(* IEC 61131-3 sources: trust-platform/examples/OSCAT/pasteurizer_quality_chain/oop/src, 3 files *)

(* ---- Main.st ---- *)
(* Record role: PasteurizerResult is a deterministic PLC-side record for tests and runtime readers. *)
TYPE PasteurizerResult :
STRUCT
    ForwardDivert : BOOL;
    DivertToRecirc : BOOL;
    RequiredTemperature : REAL;
    RequiredHoldSeconds : INT;
    SequenceStep : INT;
END_STRUCT
END_TYPE

(* Record role: QualityAlarmEvent is a deterministic PLC-side record for tests and runtime readers. *)
TYPE QualityAlarmEvent :
STRUCT
    TemperatureC : REAL;
    FlowRateLpm : REAL;
    RequiredTemperatureC : REAL;
    OperatorAck : BOOL;
    SupervisorOnline : BOOL;
END_STRUCT
END_TYPE

(* Pattern role: IQualityAlarmHandler is the contract boundary for the Chain of Responsibility and Template Method example. *)
INTERFACE IQualityAlarmHandler
    METHOD SetNext
    VAR_INPUT
        NextHandler : IQualityAlarmHandler;
    END_VAR
    END_METHOD

    METHOD Handle : BOOL
    VAR_INPUT
        Event : QualityAlarmEvent;
    END_VAR
    END_METHOD

    PROPERTY HandlerId : INT
    GET
    END_GET
    END_PROPERTY
END_INTERFACE

(* Composition role: BasePasteurizerTemplate owns the collaborating objects used by this Chain of Responsibility and Template Method example. *)
FUNCTION_BLOCK BasePasteurizerTemplate
VAR
    TempFilter : Pt2Filter;
    DivertCounter : DwordCounter;
    LastResult : PasteurizerResult;
END_VAR

METHOD PUBLIC Initialize
TempFilter.Initialize();
TempFilter.Configure(TimeConstant := T#1s, Damping := REAL#1.0, Gain := REAL#1.0);
DivertCounter.Initialize();
DivertCounter.Configure(StepSize := DWORD#1, MaxValue := DWORD#16#FFFFFFFF);
END_METHOD

METHOD PUBLIC RequiredTemperature : REAL
RequiredTemperature := REAL#72.0;
END_METHOD

METHOD PUBLIC RequiredHoldSeconds : INT
RequiredHoldSeconds := INT#15;
END_METHOD

METHOD PUBLIC Preheat : BOOL
VAR_INPUT
    ProductPresent : BOOL;
END_VAR
Preheat := ProductPresent;
END_METHOD

METHOD PUBLIC Heat : BOOL
VAR_INPUT
    ProductTemp : REAL;
END_VAR
Heat := ProductTemp >= RequiredTemperature();
END_METHOD

METHOD PUBLIC Hold : BOOL
VAR_INPUT
    HoldSeconds : INT;
END_VAR
Hold := HoldSeconds >= RequiredHoldSeconds();
END_METHOD

METHOD PUBLIC Chill : BOOL
VAR_INPUT
    FlowRate : REAL;
END_VAR
Chill := FlowRate >= REAL#100.0;
END_METHOD

METHOD PUBLIC RouteProduct : BOOL
VAR_INPUT
    HeatOk : BOOL;
    HoldOk : BOOL;
    ChillOk : BOOL;
END_VAR
RouteProduct := HeatOk AND HoldOk AND ChillOk;
END_METHOD

METHOD PUBLIC RunTemplate : PasteurizerResult
VAR_INPUT
    ProductPresent : BOOL;
    ProductTemp : REAL;
    FlowRate : REAL;
    HoldSeconds : INT;
END_VAR
VAR
    HeatOk : BOOL;
    HoldOk : BOOL;
    ChillOk : BOOL;
END_VAR
LastResult.RequiredTemperature := RequiredTemperature();
LastResult.RequiredHoldSeconds := RequiredHoldSeconds();
(* SequenceStep legend: 10=preheat wait, 20=heat, 40=recirculate/divert, 50=forward product. *)
IF NOT Preheat(ProductPresent := ProductPresent) THEN
    LastResult.SequenceStep := INT#10;
    LastResult.ForwardDivert := FALSE;
ELSIF NOT Heat(ProductTemp := ProductTemp) THEN
    LastResult.SequenceStep := INT#20;
    LastResult.ForwardDivert := FALSE;
ELSE
    HeatOk := TRUE;
    HoldOk := Hold(HoldSeconds := HoldSeconds);
    ChillOk := Chill(FlowRate := FlowRate);
    LastResult.ForwardDivert := RouteProduct(HeatOk := HeatOk, HoldOk := HoldOk, ChillOk := ChillOk);
    IF LastResult.ForwardDivert THEN
        LastResult.SequenceStep := INT#50;
    ELSE
        LastResult.SequenceStep := INT#40;
    END_IF;
END_IF;
LastResult.DivertToRecirc := NOT LastResult.ForwardDivert;
(* DwordCounter wraps COUNT_DR (edge-triggered: UP AND NOT LastUp).
   Drop the UP edge first so consecutive divert batches each generate
   a fresh rising edge and actually increment. *)
DivertCounter.Update(Up := FALSE, Down := FALSE);
IF LastResult.DivertToRecirc THEN
    DivertCounter.Update(Up := TRUE, Down := FALSE);
END_IF;
RunTemplate := LastResult;
END_METHOD
END_FUNCTION_BLOCK

(* Pattern role: MilkPasteurizer customizes inherited behavior in the Chain of Responsibility and Template Method example. *)
FUNCTION_BLOCK MilkPasteurizer EXTENDS BasePasteurizerTemplate
METHOD PUBLIC RequiredTemperature : REAL
RequiredTemperature := REAL#72.0;
END_METHOD

METHOD PUBLIC RequiredHoldSeconds : INT
RequiredHoldSeconds := INT#15;
END_METHOD
END_FUNCTION_BLOCK

(* Pattern role: CreamPasteurizer customizes inherited behavior in the Chain of Responsibility and Template Method example. *)
FUNCTION_BLOCK CreamPasteurizer EXTENDS BasePasteurizerTemplate
METHOD PUBLIC RequiredTemperature : REAL
RequiredTemperature := REAL#75.0;
END_METHOD

METHOD PUBLIC RequiredHoldSeconds : INT
RequiredHoldSeconds := INT#20;
END_METHOD
END_FUNCTION_BLOCK

(* Pattern role: LocalRecoveryHandler is a concrete implementation in the Chain of Responsibility and Template Method example. *)
FUNCTION_BLOCK LocalRecoveryHandler IMPLEMENTS IQualityAlarmHandler
VAR
    Next : IQualityAlarmHandler;
    HandlerIdValue : INT := INT#1;
    RecoveredValue : BOOL;
END_VAR

METHOD PUBLIC SetNext
VAR_INPUT
    NextHandler : IQualityAlarmHandler;
END_VAR
Next := NextHandler;
END_METHOD

METHOD PUBLIC Handle : BOOL
VAR_INPUT
    Event : QualityAlarmEvent;
END_VAR
(* Reset on entry so the flag reflects only the current event. *)
RecoveredValue := FALSE;
IF (Event.TemperatureC >= (Event.RequiredTemperatureC - REAL#1.0)) AND (Event.FlowRateLpm >= REAL#100.0) THEN
    RecoveredValue := TRUE;
    Handle := TRUE;
ELSE
    Handle := Next.Handle(Event := Event);
END_IF;
END_METHOD

METHOD PUBLIC ResetFlag
RecoveredValue := FALSE;
END_METHOD

PUBLIC PROPERTY HandlerId : INT
GET
    HandlerId := HandlerIdValue;
END_GET
END_PROPERTY

PUBLIC PROPERTY Recovered : BOOL
GET
    Recovered := RecoveredValue;
END_GET
END_PROPERTY
END_FUNCTION_BLOCK

(* Pattern role: OperatorAcknowledgeHandler is a concrete implementation in the Chain of Responsibility and Template Method example. *)
FUNCTION_BLOCK OperatorAcknowledgeHandler IMPLEMENTS IQualityAlarmHandler
VAR
    Next : IQualityAlarmHandler;
    HandlerIdValue : INT := INT#2;
    AcknowledgedValue : BOOL;
END_VAR

METHOD PUBLIC SetNext
VAR_INPUT
    NextHandler : IQualityAlarmHandler;
END_VAR
Next := NextHandler;
END_METHOD

METHOD PUBLIC Handle : BOOL
VAR_INPUT
    Event : QualityAlarmEvent;
END_VAR
(* Reset on entry so the flag reflects only the current event. *)
AcknowledgedValue := FALSE;
IF Event.OperatorAck THEN
    AcknowledgedValue := TRUE;
    Handle := TRUE;
ELSE
    Handle := Next.Handle(Event := Event);
END_IF;
END_METHOD

METHOD PUBLIC ResetFlag
AcknowledgedValue := FALSE;
END_METHOD

PUBLIC PROPERTY HandlerId : INT
GET
    HandlerId := HandlerIdValue;
END_GET
END_PROPERTY

PUBLIC PROPERTY Acknowledged : BOOL
GET
    Acknowledged := AcknowledgedValue;
END_GET
END_PROPERTY
END_FUNCTION_BLOCK

(* Pattern role: SupervisorEscalateHandler is a concrete implementation in the Chain of Responsibility and Template Method example. *)
FUNCTION_BLOCK SupervisorEscalateHandler IMPLEMENTS IQualityAlarmHandler
VAR
    Next : IQualityAlarmHandler;
    HandlerIdValue : INT := INT#3;
    EscalatedValue : BOOL;
END_VAR

METHOD PUBLIC SetNext
VAR_INPUT
    NextHandler : IQualityAlarmHandler;
END_VAR
Next := NextHandler;
END_METHOD

METHOD PUBLIC Handle : BOOL
VAR_INPUT
    Event : QualityAlarmEvent;
END_VAR
(* Reset on entry so the flag reflects only the current event. *)
EscalatedValue := FALSE;
IF Event.SupervisorOnline THEN
    EscalatedValue := TRUE;
    Handle := TRUE;
ELSE
    Handle := Next.Handle(Event := Event);
END_IF;
END_METHOD

METHOD PUBLIC ResetFlag
EscalatedValue := FALSE;
END_METHOD

PUBLIC PROPERTY HandlerId : INT
GET
    HandlerId := HandlerIdValue;
END_GET
END_PROPERTY

PUBLIC PROPERTY Escalated : BOOL
GET
    Escalated := EscalatedValue;
END_GET
END_PROPERTY
END_FUNCTION_BLOCK

(* Pattern role: BatchAbortHandler is a concrete implementation in the Chain of Responsibility and Template Method example. *)
FUNCTION_BLOCK BatchAbortHandler IMPLEMENTS IQualityAlarmHandler
VAR
    HandlerIdValue : INT := INT#4;
    AbortedValue : BOOL;
END_VAR

METHOD PUBLIC SetNext
VAR_INPUT
    NextHandler : IQualityAlarmHandler;
END_VAR
END_METHOD

METHOD PUBLIC Handle : BOOL
VAR_INPUT
    Event : QualityAlarmEvent;
END_VAR
(* Last handler in chain: always handles. Flag is set fresh each call. *)
AbortedValue := TRUE;
Handle := TRUE;
END_METHOD

METHOD PUBLIC ResetFlag
AbortedValue := FALSE;
END_METHOD

PUBLIC PROPERTY HandlerId : INT
GET
    HandlerId := HandlerIdValue;
END_GET
END_PROPERTY

PUBLIC PROPERTY Aborted : BOOL
GET
    Aborted := AbortedValue;
END_GET
END_PROPERTY
END_FUNCTION_BLOCK

(* Composition role: PasteurizerController owns the collaborating objects used by this Chain of Responsibility and Template Method example. *)
FUNCTION_BLOCK PasteurizerController
VAR
    Milk : MilkPasteurizer;
    Cream : CreamPasteurizer;
    Local : LocalRecoveryHandler;
    Operator : OperatorAcknowledgeHandler;
    Supervisor : SupervisorEscalateHandler;
    Abort : BatchAbortHandler;
    AlarmChain : IQualityAlarmHandler;
    LastResultValue : PasteurizerResult;
    LastHandlerIdValue : INT;
END_VAR

METHOD PUBLIC Initialize
Milk.Initialize();
Cream.Initialize();
Local.SetNext(NextHandler := Operator);
Operator.SetNext(NextHandler := Supervisor);
Supervisor.SetNext(NextHandler := Abort);
AlarmChain := Local;
END_METHOD

METHOD PUBLIC Update : PasteurizerResult
VAR_INPUT
    RecipeId : INT;
    ProductTemp : REAL;
    FlowRate : REAL;
    HoldSeconds : INT;
    OperatorAck : BOOL;
    SupervisorOnline : BOOL;
END_VAR
VAR
    Event : QualityAlarmEvent;
END_VAR
(* Clear cross-batch sticky state so LastHandlerId reflects only the current batch. *)
LastHandlerIdValue := INT#0;
Local.ResetFlag();
Operator.ResetFlag();
Supervisor.ResetFlag();
Abort.ResetFlag();
IF RecipeId = INT#2 THEN
    LastResultValue := Cream.RunTemplate(ProductPresent := TRUE, ProductTemp := ProductTemp, FlowRate := FlowRate, HoldSeconds := HoldSeconds);
ELSE
    LastResultValue := Milk.RunTemplate(ProductPresent := TRUE, ProductTemp := ProductTemp, FlowRate := FlowRate, HoldSeconds := HoldSeconds);
END_IF;

IF LastResultValue.DivertToRecirc THEN
    Event.TemperatureC := ProductTemp;
    Event.FlowRateLpm := FlowRate;
    Event.RequiredTemperatureC := LastResultValue.RequiredTemperature;
    Event.OperatorAck := OperatorAck;
    Event.SupervisorOnline := SupervisorOnline;
    AlarmChain.Handle(Event := Event);
    IF Abort.Aborted THEN
        LastHandlerIdValue := Abort.HandlerId;
    ELSIF Supervisor.Escalated THEN
        LastHandlerIdValue := Supervisor.HandlerId;
    ELSIF Operator.Acknowledged THEN
        LastHandlerIdValue := Operator.HandlerId;
    ELSIF Local.Recovered THEN
        LastHandlerIdValue := Local.HandlerId;
    END_IF;
END_IF;
Update := LastResultValue;
END_METHOD

PUBLIC PROPERTY ForwardDivert : BOOL
GET
    ForwardDivert := LastResultValue.ForwardDivert;
END_GET
END_PROPERTY

PUBLIC PROPERTY BatchAborted : BOOL
GET
    BatchAborted := Abort.Aborted;
END_GET
END_PROPERTY

PUBLIC PROPERTY LastHandlerId : INT
GET
    LastHandlerId := LastHandlerIdValue;
END_GET
END_PROPERTY

PUBLIC PROPERTY RequiredTemperature : REAL
GET
    RequiredTemperature := LastResultValue.RequiredTemperature;
END_GET
END_PROPERTY
END_FUNCTION_BLOCK

(* Scan role: Main wires the example objects and exposes the PLC call path under test. *)
PROGRAM Main
VAR
    Pasteurizer : PasteurizerController;
    RecipeId : INT;
    ProductTempRaw : INT;
    FlowRateRaw : INT;
    OperatorAck : BOOL;
    SupervisorOnline : BOOL;
    Result : PasteurizerResult;
    ForwardValveOut : BOOL;
    DivertValveOut : BOOL;
    AlarmOut : BOOL;
END_VAR

Pasteurizer.Initialize();
Result := Pasteurizer.Update(RecipeId := RecipeId, ProductTemp := INT_TO_REAL(ProductTempRaw), FlowRate := INT_TO_REAL(FlowRateRaw), HoldSeconds := INT#15, OperatorAck := OperatorAck, SupervisorOnline := SupervisorOnline);
ForwardValveOut := Result.ForwardDivert;
DivertValveOut := Result.DivertToRecirc;
AlarmOut := Result.DivertToRecirc;
END_PROGRAM

(* ---- Configuration.st ---- *)
CONFIGURATION PasteurizerQualityChainOopConfiguration
RESOURCE Cpu0 ON PLC
    TASK MainTask (INTERVAL := T#100ms, PRIORITY := 1);
    PROGRAM Pasteurizer WITH MainTask : Main;
END_RESOURCE
VAR_CONFIG
    Pasteurizer.RecipeId AT %IW0 : INT;
    Pasteurizer.ProductTempRaw AT %IW2 : INT;
    Pasteurizer.FlowRateRaw AT %IW4 : INT;
    Pasteurizer.OperatorAck AT %IX0.0 : BOOL;
    Pasteurizer.SupervisorOnline AT %IX0.1 : BOOL;
    Pasteurizer.ForwardValveOut AT %QX0.0 : BOOL;
    Pasteurizer.DivertValveOut AT %QX0.1 : BOOL;
    Pasteurizer.AlarmOut AT %QX0.2 : BOOL;
END_VAR
END_CONFIGURATION

(* ---- Tests.st ---- *)
TEST_PROGRAM PasteurizerTemplateUsesRecipeHooks
VAR
    Milk : MilkPasteurizer;
    Cream : CreamPasteurizer;
    MilkResult : PasteurizerResult;
    CreamResult : PasteurizerResult;
END_VAR

Milk.Initialize();
Cream.Initialize();
MilkResult := Milk.RunTemplate(ProductPresent := TRUE, ProductTemp := REAL#73.0, FlowRate := REAL#120.0, HoldSeconds := INT#15);
CreamResult := Cream.RunTemplate(ProductPresent := TRUE, ProductTemp := REAL#73.0, FlowRate := REAL#120.0, HoldSeconds := INT#15);
ASSERT_TRUE(IN := MilkResult.ForwardDivert);
ASSERT_FALSE(IN := CreamResult.ForwardDivert);
ASSERT_NEAR(EXPECTED := REAL#75.0, ACTUAL := CreamResult.RequiredTemperature, DELTA := REAL#0.001);
ASSERT_EQUAL(EXPECTED := INT#20, ACTUAL := CreamResult.RequiredHoldSeconds);
END_TEST_PROGRAM

TEST_PROGRAM QualityAlarmChainEscalatesToAbortWhenUnhandled
VAR
    Controller : PasteurizerController;
    Result : PasteurizerResult;
END_VAR

Controller.Initialize();
Result := Controller.Update(RecipeId := INT#1, ProductTemp := REAL#68.0, FlowRate := REAL#90.0, HoldSeconds := INT#5, OperatorAck := FALSE, SupervisorOnline := FALSE);
ASSERT_FALSE(IN := Result.ForwardDivert);
ASSERT_TRUE(IN := Controller.BatchAborted);
ASSERT_EQUAL(EXPECTED := INT#4, ACTUAL := Controller.LastHandlerId);
END_TEST_PROGRAM

TEST_PROGRAM QualityAlarmChainStopsAtOperatorAcknowledge
VAR
    Controller : PasteurizerController;
    Result : PasteurizerResult;
END_VAR

Controller.Initialize();
Result := Controller.Update(RecipeId := INT#1, ProductTemp := REAL#68.0, FlowRate := REAL#90.0, HoldSeconds := INT#5, OperatorAck := TRUE, SupervisorOnline := FALSE);
ASSERT_FALSE(IN := Result.ForwardDivert);
ASSERT_FALSE(IN := Controller.BatchAborted);
ASSERT_EQUAL(EXPECTED := INT#2, ACTUAL := Controller.LastHandlerId);
END_TEST_PROGRAM

(* Multi-batch chain regression: drives several different batches
   through one Controller. Catches the same bug class as
   tunnel_washer_chain — handler flags or LastHandlerId leaking
   between events because handlers don't reset their per-call state. *)
TEST_PROGRAM PasteurizerChainHandlesMultipleBatchesIndependently
VAR
    Controller : PasteurizerController;
    Result : PasteurizerResult;
END_VAR

Controller.Initialize();

(* Batch 1: bad temp + supervisor online -> escalates to supervisor (3) *)
Result := Controller.Update(RecipeId := INT#1, ProductTemp := REAL#68.0, FlowRate := REAL#90.0, HoldSeconds := INT#5, OperatorAck := FALSE, SupervisorOnline := TRUE);
ASSERT_EQUAL(EXPECTED := INT#3, ACTUAL := Controller.LastHandlerId);

(* Batch 2: same bad temp but operator now acks -> stops at handler 2.
   LastHandlerId must reflect the new outcome, not the previous (3). *)
Result := Controller.Update(RecipeId := INT#1, ProductTemp := REAL#68.0, FlowRate := REAL#90.0, HoldSeconds := INT#5, OperatorAck := TRUE, SupervisorOnline := FALSE);
ASSERT_EQUAL(EXPECTED := INT#2, ACTUAL := Controller.LastHandlerId);

(* Batch 3: nothing helps -> escalates to abort (4) *)
Result := Controller.Update(RecipeId := INT#1, ProductTemp := REAL#68.0, FlowRate := REAL#90.0, HoldSeconds := INT#5, OperatorAck := FALSE, SupervisorOnline := FALSE);
ASSERT_EQUAL(EXPECTED := INT#4, ACTUAL := Controller.LastHandlerId);
ASSERT_TRUE(IN := Controller.BatchAborted);
END_TEST_PROGRAM

(* Happy path: in-spec batch forwards directly. *)
TEST_PROGRAM PasteurizerForwardsInSpecBatchWithoutEscalation
VAR
    Controller : PasteurizerController;
    Result : PasteurizerResult;
END_VAR
Controller.Initialize();
Result := Controller.Update(RecipeId := INT#1, ProductTemp := REAL#74.0, FlowRate := REAL#120.0, HoldSeconds := INT#16, OperatorAck := FALSE, SupervisorOnline := FALSE);
ASSERT_TRUE(IN := Result.ForwardDivert);
ASSERT_FALSE(IN := Controller.BatchAborted);
END_TEST_PROGRAM

(* LocalRecoveryHandler in isolation: requires temp within 1 C AND flow >= 100. *)
TEST_PROGRAM LocalRecoveryHandlerHandlesNearMissOnly
VAR
    Local : LocalRecoveryHandler;
    Terminal : BatchAbortHandler;
    Event : QualityAlarmEvent;
END_VAR
Local.SetNext(NextHandler := Terminal);

(* Within 1 C of required + flow ok: handles *)
Event.RequiredTemperatureC := REAL#73.0;
Event.TemperatureC := REAL#72.5;
Event.FlowRateLpm := REAL#110.0;
Event.OperatorAck := FALSE;
Event.SupervisorOnline := FALSE;
Local.Handle(Event := Event);
ASSERT_TRUE(IN := Local.Recovered);

(* Temp too far below required: passes through *)
Event.TemperatureC := REAL#68.0;
Local.Handle(Event := Event);
ASSERT_FALSE(IN := Local.Recovered);

(* Temp ok but flow too low: passes through *)
Event.TemperatureC := REAL#72.5;
Event.FlowRateLpm := REAL#90.0;
Local.Handle(Event := Event);
ASSERT_FALSE(IN := Local.Recovered);

(* Boundary: flow exactly 100 - inclusive *)
Event.FlowRateLpm := REAL#100.0;
Local.Handle(Event := Event);
ASSERT_TRUE(IN := Local.Recovered);

(* Boundary: temp exactly Required - 1.0 - inclusive *)
Event.TemperatureC := REAL#72.0;
Event.FlowRateLpm := REAL#100.0;
Local.Handle(Event := Event);
ASSERT_TRUE(IN := Local.Recovered);
END_TEST_PROGRAM

(* OperatorAcknowledgeHandler isolation. *)
TEST_PROGRAM OperatorAcknowledgeHandlerHandlesOnlyWhenAckPresent
VAR
    Operator : OperatorAcknowledgeHandler;
    Terminal : BatchAbortHandler;
    Event : QualityAlarmEvent;
END_VAR
Operator.SetNext(NextHandler := Terminal);

Event.OperatorAck := TRUE;
Operator.Handle(Event := Event);
ASSERT_TRUE(IN := Operator.Acknowledged);

Event.OperatorAck := FALSE;
Operator.Handle(Event := Event);
ASSERT_FALSE(IN := Operator.Acknowledged);
END_TEST_PROGRAM

(* SupervisorEscalateHandler isolation. *)
TEST_PROGRAM SupervisorEscalateHandlerHandlesOnlyWhenSupervisorOnline
VAR
    Supervisor : SupervisorEscalateHandler;
    Terminal : BatchAbortHandler;
    Event : QualityAlarmEvent;
END_VAR
Supervisor.SetNext(NextHandler := Terminal);

Event.SupervisorOnline := TRUE;
Supervisor.Handle(Event := Event);
ASSERT_TRUE(IN := Supervisor.Escalated);

Event.SupervisorOnline := FALSE;
Supervisor.Handle(Event := Event);
ASSERT_FALSE(IN := Supervisor.Escalated);
END_TEST_PROGRAM

(* Local recovery is preferred over operator/supervisor when both could handle. *)
TEST_PROGRAM PasteurizerChainPrefersLocalRecoveryWhenEligible
VAR
    Controller : PasteurizerController;
    Result : PasteurizerResult;
END_VAR
Controller.Initialize();
(* Slightly-off temp (below milk required 72 C) + flow >= 100 + operator
   + supervisor all available. Heat fails so divert triggers and chain
   runs. Order Local -> Operator -> Supervisor -> Abort. Local wins
   because TemperatureC (71.5) >= RequiredTemperatureC - 1.0 (71.0)
   and FlowRateLpm (110) >= 100.0. *)
Result := Controller.Update(RecipeId := INT#1, ProductTemp := REAL#71.5, FlowRate := REAL#110.0, HoldSeconds := INT#16, OperatorAck := TRUE, SupervisorOnline := TRUE);
ASSERT_FALSE(IN := Result.ForwardDivert);
ASSERT_EQUAL(EXPECTED := INT#1, ACTUAL := Controller.LastHandlerId);
END_TEST_PROGRAM

(* Recipe variant difference: cream requires 75 C, milk requires 73 C. *)
TEST_PROGRAM PasteurizerCreamRecipeRequiresHigherTemperature
VAR
    Controller : PasteurizerController;
    Result : PasteurizerResult;
END_VAR
Controller.Initialize();

(* 73 C: fine for milk (recipe 1), insufficient for cream (recipe 2) *)
Result := Controller.Update(RecipeId := INT#1, ProductTemp := REAL#73.0, FlowRate := REAL#120.0, HoldSeconds := INT#15, OperatorAck := FALSE, SupervisorOnline := FALSE);
ASSERT_TRUE(IN := Result.ForwardDivert);

(* Cream needs 75 - 73 falls into LocalRecovery range only with hold *)
Result := Controller.Update(RecipeId := INT#2, ProductTemp := REAL#73.0, FlowRate := REAL#120.0, HoldSeconds := INT#15, OperatorAck := FALSE, SupervisorOnline := FALSE);
ASSERT_FALSE(IN := Result.ForwardDivert);

(* 75 C: cream passes *)
Result := Controller.Update(RecipeId := INT#2, ProductTemp := REAL#76.0, FlowRate := REAL#120.0, HoldSeconds := INT#20, OperatorAck := FALSE, SupervisorOnline := FALSE);
ASSERT_TRUE(IN := Result.ForwardDivert);
END_TEST_PROGRAM
